// TIA Portal V20 export
Screen "Call_ServiceButtons_2"  1276x673
  ScreenItem "Title_OPMode1_ScreenOverview_X390_Y2" at 5,7 size 1262x30  Type=HmiTextBox
  ScreenItem "Faceplate container_5" at 0,33 size 622x206  Type=HmiFaceplateContainer
  ScreenItem "Text box_5" at 0,0 size 622x30  Type=HmiTextBox
  ScreenItem "Faceplate container_7" at 0,33 size 622x206  Type=HmiFaceplateContainer
  ScreenItem "Text box_7" at 0,0 size 622x30  Type=HmiTextBox
  ScreenItem "Faceplate container_8" at 0,33 size 622x206  Type=HmiFaceplateContainer
  ScreenItem "Text box_8" at 0,0 size 622x30  Type=HmiTextBox
  ScreenItem "Faceplate container_6" at 5,73 size 619x179  Type=HmiFaceplateContainer
  ScreenItem "Text box_6" at 5,40 size 622x30  Type=HmiTextBox
  ScreenItem "Faceplate container_9" at 645,73 size 619x179  Type=HmiFaceplateContainer
  ScreenItem "Text box_9" at 644,40 size 622x30  Type=HmiTextBox
